SUBAPPLICATION SubApp_PC_A (* Geraet A: Flip-Flop (opcua.adoc): SUBSCRIBE Flip -> E_SWITCH/E_SR -> PUBLISH Flop; Input_I1 schreibt Flip, Output_Q1 zeigt Flop (= NICHT I1) *)
  (* Standard: 61499-2; Description: Copyright (c) 2026 Meisterschulen am Ostbahnhof This program and the accompanying materials are made available under the terms of the Eclipse Public License 2.0 which is available at https://www.eclipse.org/legal/epl-2.0/ SPDX-License-Identifier: EPL-2.0 *)
  (* Version 1.0, 2026-10-18, Franz Höpfinger, Meisterschulen am Ostbahnhof, opcua.adoc-Beispiel auf zwei Geraeten *)
  PACKAGE subapp::Training_13_OPC_UA_RES;
  IMPORT VV::const::OPC_UA::myOpcUaAddresses::T13_FLIP_REMOTE_WRITE;
  IMPORT VV::const::OPC_UA::myOpcUaAddresses::T13_FLOP_REMOTE_SUBSCRIBE;
  IMPORT logiBUS::io::DI::logiBUS_DI::Input_I1;
  IMPORT logiBUS::io::DQ::logiBUS_DO::Output_Q1;
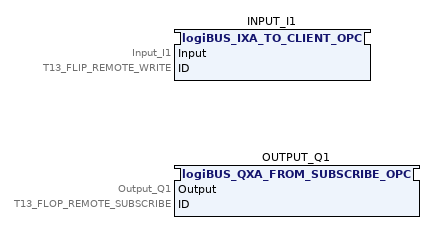
  SUBAPPS
    INPUT_I1 : MyLib::sys::logiBUS_IXA_TO_CLIENT_OPC(Input := Input_I1, ID := T13_FLIP_REMOTE_WRITE);
    OUTPUT_Q1 : MyLib::sys::logiBUS_QXA_FROM_SUBSCRIBE_OPC(Output := Output_Q1, ID := T13_FLOP_REMOTE_SUBSCRIBE);
  END_SUBAPPS
END_SUBAPPLICATION
